(* IEC 61131-3 sources: rusty/tests/lit/single/actions, 5 files *)

(* ---- action_call_with_var_in_out.st ---- *)
// RUN: %COMPILE %s && %RUN | %CHECK %s
// Regression coverage for #1576 (fixed in commit 2b3388f). Calling an action
// that inherits a `VAR_IN_OUT` parameter from its parent FB must store the
// caller's address into the FB's in-out slot before invoking the action.
// Before the fix the slot stayed NULL — the action then dereferenced a null
// pointer and segfaulted at runtime.

PROGRAM mainProg
VAR
    fb : fb_t;
    localBool : BOOL;
END_VAR
    localBool := TRUE;
    fb.foo(myInOut := localBool);

    localBool := FALSE;
    fb.foo(myInOut := localBool);
END_PROGRAM

FUNCTION_BLOCK fb_t
VAR_IN_OUT
    myInOut : BOOL;
END_VAR
END_FUNCTION_BLOCK

ACTIONS
    ACTION foo
        // CHECK: myInout = 1
        // CHECK: myInout = 0
        printf('myInout = %d$N', myInOut);
    END_ACTION
END_ACTIONS

FUNCTION main : DINT
    mainProg();
    main := 0;
END_FUNCTION

(* ---- for_loop_in_action.st ---- *)
// RUN: %COMPILE %s && %RUN | %CHECK %s
// Regression: a FOR loop inside an action must resolve its desugared temporaries (#1784).

PROGRAM mainProg
VAR
    acc : DINT;
    i : DINT;
END_VAR
    foo();
END_PROGRAM

ACTIONS
    ACTION foo
        acc := 0;
        FOR i := 1 TO 10 DO
            acc := acc + i;
        END_FOR
        printf('for=%d$N', acc); // CHECK: for=55
    END_ACTION
END_ACTIONS

FUNCTION main : DINT
    mainProg();
    main := 0;
END_FUNCTION

(* ---- nested_loops_in_action.st ---- *)
// RUN: %COMPILE %s && %RUN | %CHECK %s
// Regression: nested loops inside an action must re-initialize their inner temporaries (#1784).

PROGRAM mainProg
VAR
    acc : DINT;
    i : DINT;
    j : DINT;
END_VAR
    foo();
END_PROGRAM

ACTIONS
    ACTION foo
        acc := 0;
        FOR i := 1 TO 3 DO
            FOR j := 1 TO 3 DO
                acc := acc + 1;
            END_FOR
        END_FOR
        printf('nested=%d$N', acc); // CHECK: nested=9
    END_ACTION
END_ACTIONS

FUNCTION main : DINT
    mainProg();
    main := 0;
END_FUNCTION

(* ---- repeat_loop_in_action.st ---- *)
// RUN: %COMPILE %s && %RUN | %CHECK %s
// Regression: a REPEAT loop inside an action must resolve its `__ran_once_*` temporary (#1784).

PROGRAM mainProg
VAR
    acc : DINT;
END_VAR
    foo();
END_PROGRAM

ACTIONS
    ACTION foo
        acc := 0;
        REPEAT
            acc := acc + 1;
        UNTIL acc >= 3
        END_REPEAT
        printf('repeat=%d$N', acc); // CHECK: repeat=3
    END_ACTION
END_ACTIONS

FUNCTION main : DINT
    mainProg();
    main := 0;
END_FUNCTION

(* ---- while_loop_in_action.st ---- *)
// RUN: %COMPILE %s && %RUN | %CHECK %s
// Regression: a WHILE loop inside an action must resolve against the parent POU's members (#1784).

PROGRAM mainProg
VAR
    acc : DINT;
    i : DINT;
END_VAR
    foo();
END_PROGRAM

ACTIONS
    ACTION foo
        acc := 0;
        i := 0;
        WHILE i < 5 DO
            acc := acc + 1;
            i := i + 1;
        END_WHILE
        printf('while=%d$N', acc); // CHECK: while=5
    END_ACTION
END_ACTIONS

FUNCTION main : DINT
    mainProg();
    main := 0;
END_FUNCTION
